TYPE ST_DiagnosticElementOut :
STRUCT
    sName: STRING(20) := 'Unnamed';
    sAlarmMsg: STRING(20) := 'Not defined';
    bRun: BOOL;
    bReady: BOOL;
    bSafe: BOOL;
    bError: BOOL;
    bCycle: BOOL;
    bReset: BOOL;
END_STRUCT
END_TYPE

(* stored: Version 1.1.0.1
   DUT ST_DiagnosticElementOut: Id {a03f9acf-2cc9-020d-31d2-8b63b6993c66} *)
